(* IEC 61131-3 sources: codesys-to-s7/tests/corpus/C2S7-GFX-GOTO/pos, 1 file *)

(* ---- input.st ---- *)
FUNCTION_BLOCK FB_J
VAR_INPUT
    a : BOOL;
END_VAR
VAR
    i : INT;
END_VAR
IF a THEN
    JMP lbl;
END_IF
i := 1;
lbl:
i := i + 2;
END_FUNCTION_BLOCK
